(* PLC project v0.5.4_.project, CODESYS CODESYS V3.5 SP19 Patch 1 *)
(* stored: creationDateTime 2026-08-04T04:31:53.0000133, modificationDateTime 2026-08-04T04:31:03.5723483 *)

PROGRAM PRG_Oracle_Nested
  VAR
    instSafety : FB_Safety_EmergencyManagement;  (* ou tout FB avec output struct *)
    ArmingSeqStep : INT;
    PowerKeepAlive_A_RQ : BOOL;
  END_VAR

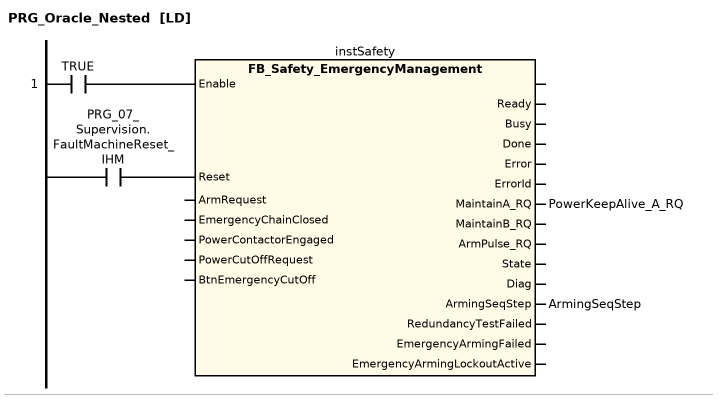
(* LD diagram, written out as Structured Text *)

instSafety(Enable := TRUE, Reset := PRG_07_Supervision.FaultMachineReset_IHM, ArmRequest := , EmergencyChainClosed := , PowerContactorEngaged := , PowerCutOffRequest := , BtnEmergencyCutOff := , MaintainA_RQ => PowerKeepAlive_A_RQ, ArmingSeqStep => ArmingSeqStep);
END_PROGRAM
